Fanuc KAREL source: KD00065.KL

PROGRAM KD00065
%NOLOCKGROUP
VAR
  I: INTEGER
  J: INTEGER
  B: BOOLEAN
  R: REAL
  S: STRING[80]
BEGIN
  CONDITION[1]:
  WHEN DIN[1] = ON DO
    NOABORT
  ENDCONDITION
END KD00065
